FUNCTION_BLOCK MOD_StateView (* Tells the block it sits in the module's PackML state, and asks for it once at start. Technical: The module's PackML state from its local channel; asks for the current value at INIT *)
  (* Standard: 61499-2 *)
  (* Version 0.1, 2026-09-28, Project contributors, AAU Smart Production Lab *)
  PACKAGE modlib;
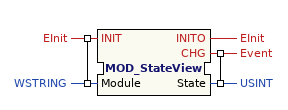
  EVENT_INPUT
    INIT : EInit WITH Module; (* Initialise, once at start-up (the INIT chain); takes the values given with it *)
  END_EVENT
  EVENT_OUTPUT
    INITO : EInit; (* Initialised: the next block of the INIT chain goes on *)
    CHG WITH State; (* The value changed *)
  END_EVENT
  VAR_INPUT
    Module : WSTRING; (* The module's name; its local channels are named after it (loc[<Module>/...]) *)
  END_VAR
  VAR_OUTPUT
    State : USINT; (* PackML state: 1 Clearing, 2 Stopped, 3 Starting, 4 Idle, 6 Execute, 7 Stopping, 8 Aborting, 9 Aborted, 15 Resetting *)
  END_VAR
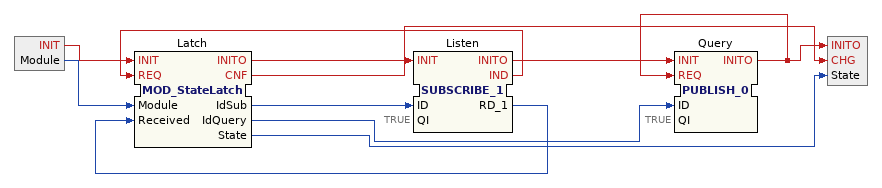
  FBS
    Latch : modlib::MOD_StateLatch; (* Keeps the last module state heard. *)
    Listen : iec61499::net::SUBSCRIBE_1(QI := TRUE); (* Listens to the module's state channel. *)
    Query : iec61499::net::PUBLISH_0(QI := TRUE); (* Asks for the state once at start. *)
  END_FBS
  EVENT_CONNECTIONS
    INIT TO Latch.INIT;
    Latch.INITO TO Listen.INIT;
    Listen.INITO TO Query.INIT;
    Query.INITO TO Query.REQ;
    Query.INITO TO INITO;
    Listen.IND TO Latch.REQ;
    Latch.CNF TO CHG;
  END_CONNECTIONS
  DATA_CONNECTIONS
    Module TO Latch.Module;
    Latch.IdSub TO Listen.ID;
    Latch.IdQuery TO Query.ID;
    Listen.RD_1 TO Latch.Received;
    Latch.State TO State;
  END_CONNECTIONS
END_FUNCTION_BLOCK
